FUNCTION_BLOCK FB_MotorFake IMPLEMENTS I_Motor
VAR_INPUT
    fault : BOOL;
END_VAR
VAR_OUTPUT
    updates : UDINT;
END_VAR
VAR
    speed : LREAL := 0.5;
    runningState : BOOL;
END_VAR

(* Update is called through I_Motor by the conveyor. *)

METHOD PUBLIC Update
VAR_INPUT
    run : BOOL;
    delay : TIME;
END_VAR
VAR_INST
    startup : TON;
END_VAR
updates := updates + 1;
startup(IN := run AND NOT fault, PT := delay);
THIS^.runningState := startup.Q;
END_METHOD

PROPERTY PUBLIC SpeedSetpoint : LREAL
GET
SpeedSetpoint := THIS^.speed;
END_GET
SET
THIS^.speed := LIMIT(0.0, SpeedSetpoint, 1.0);
END_SET
END_PROPERTY

PROPERTY PUBLIC Running : BOOL
GET
Running := THIS^.runningState;
END_GET
END_PROPERTY

PROPERTY PUBLIC Faulted : BOOL
GET
Faulted := fault;
END_GET
END_PROPERTY

PROPERTY PUBLIC ActualSpeed : LREAL
GET
IF THIS^.runningState THEN
    ActualSpeed := THIS^.speed;
ELSE
    ActualSpeed := 0.0;
END_IF;
END_GET
END_PROPERTY

END_FUNCTION_BLOCK

(* stored: Version 1.1.0.1, ProductVersion 3.1 *)
